FUNCTION_BLOCK HighLevelAlarmFB
  VAR
  END_VAR
  VAR_INPUT
    AtOrAbove75 : BOOL;
  END_VAR
  VAR_OUTPUT
    Alarm : BOOL;
  END_VAR

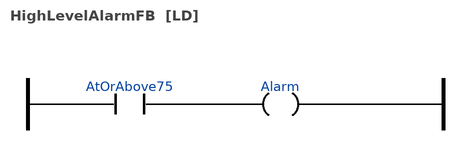
(* LD diagram, written out as Structured Text *)
Alarm := AtOrAbove75;
END_FUNCTION_BLOCK
